TYPE ET_BOSCH_Reset :
(
	eWaitExecute := 0,
	eInit,
	eReadDriveError,
	eWriteResetDriver,
	eEraseResetDriver,
	eChMCReset,
	eMCReset,
	eWfMCReset,
	eDone := 197,
	eError := 198,
	eNotExecute := 199
);
END_TYPE

(* stored: Version 1.1.0.1, ProductVersion 3.1.4024.15
   DUT ET_BOSCH_Reset: Id {649d533f-5203-4215-bf4d-d6b4744fb2f8} *)
